Staubli VAL3: safeCheck.dtx

mdesc mNomSpeed
num nToolIndex
public num nIO_Zoneindex[16]
public num nIO_spindex[16]
public dio O_safePoint[16]
public dio O_safeZone
